Fanuc KAREL source: ka00227.KL

-- PROVISIONAL review KL for V770-1; original PC SHA256 86a8d20ac60d94240d314fae7cd35b76fbb97bb579a6cb9599f9cfa7ec9d4621
-- Incomplete behavior may be omitted. Consult companion uncertainty JSON. Do not deploy.
PROGRAM KA00227
%NOLOCKGROUP
-- UNRESOLVED_DECL SRC type=001100
-- UNRESOLVED_DECL DST type=001100
BEGIN
  -- UNRESOLVED_PC offsets 5-20; opcodes 22,22,30
  -- UNRESOLVED_PC offsets 25-29; opcodes 7F
END KA00227
